TYPE TcoKukaKss_Inputs_v_9_3_x :
STRUCT
	Inputs AT %I* : ARRAY[0..63] OF BYTE;
END_STRUCT
END_TYPE

(* stored: Version 1.1.0.1, ProductVersion 3.1.4024.12
   DUT TcoKukaKss_Inputs_v_9_3_x: Id {b3d8b24e-bc0a-4500-80a0-475f0be18b8b} *)
